Fanuc KAREL source: kb00042.KL

-- PROVISIONAL review KL for V1013-1; original PC SHA256 d386b1236b1dd349aff5aa945dc56c551ec6e3072338aea83454c981870ad6a5
-- Incomplete behavior may be omitted. Consult companion uncertainty JSON. Do not deploy.
PROGRAM KB00042
%NOLOCKGROUP
BEGIN
  -- UNRESOLVED_PC offsets 5-14; opcodes 3F,75
  -- UNRESOLVED_PC offsets 19-26; opcodes 9D,23
  -- UNRESOLVED_PC offsets 31-49; opcodes 27,22,2A,22,31
  -- UNRESOLVED_PC offsets 54-58; opcodes 7F
END KB00042
